# EPICS substitutions: db/Beckhoff_7XXX/ecmcEX72XX_OPT_torqueOffset.substitutions
file "ecmc_analogOutput-chX.template"
{
  pattern {CH_ID, sourceName, KEY, suffix, DESC, EGU, ESLO, PREC, LOPR, HOPR, LOLO, LOW, HIGH, HIHI, HYST, LLSV, LSV, HSV, HHSV}
          {"$(OPT_CH_ID=01)", "torqueOffset", "Drv", "-TrqOff", "Torque Offset", "%", 0.1, 1, -200, 200, 0, 0, 0, 0, 0, "NO_ALARM", "NO_ALARM", "NO_ALARM", "NO_ALARM"}
}
